Yaskawa INFORM job: 1B.JBI

/JOB
//NAME 1B
//POS
///NPOS 156,156,156,0,0,0
///TOOL 0
///POSTYPE PULSE
///PULSE
C00000=-283,-101162,-84213,3710,-80188,-1936
C00001=-283,-101162,-84213,3710,-80188,-1936
C00002=122740,19157,4035,6182,-38864,-3236
C00003=113896,2387,-35230,-12259,-73873,84724
C00004=118077,18356,-38305,-5593,-67110,82106
C00005=118077,18356,-38305,-5593,-67110,82106
C00006=124954,18047,-39669,933,-60764,50503
C00007=142043,41533,-31174,35083,-70402,26464
C00008=142043,41533,-31174,35083,-70402,26464
C00009=142043,41533,-31174,35083,-70402,26464
C00010=138380,29006,-36364,33085,-57919,16054
C00011=120169,44405,-13547,1008,-67670,-3095
C00012=105097,34464,-28801,-23051,-62948,-22596
C00013=95890,29559,-44356,-45908,-59845,-13171
C00014=95890,29559,-44356,-45908,-59845,-13171
C00015=95890,29559,-44356,-45908,-59845,-13171
C00016=100253,12469,-52865,-35215,-53568,-35172
C00017=118532,18556,-38083,-5671,-67115,-85546
C00018=114163,-2238,-37790,-11674,-74104,-76880
C00019=113860,-11716,-39905,-11456,-77647,88229
C00020=114263,6764,-46011,-12423,-64616,86905
C00021=114386,12590,-43965,-12584,-62907,81236
C00022=114386,12590,-43965,-12584,-62907,81236
C00023=125315,10262,-47133,583,-53482,49755
C00024=142444,42695,-30785,35929,-71152,26137
C00025=142444,42695,-30785,35929,-71152,26137
C00026=142444,42695,-30785,35929,-71152,26137
C00027=138388,28635,-37117,33161,-57685,15974
C00028=120215,45689,-12379,963,-68675,-3097
C00029=105043,34518,-28884,-23053,-62885,-22568
C00030=94945,31173,-44363,-48216,-61083,-12269
C00031=94945,31173,-44363,-48216,-61083,-12269
C00032=94945,31173,-44363,-48216,-61083,-12269
C00033=98921,36729,-33454,-32527,-73118,-41437
C00034=120115,8294,-47151,319,-58957,-81109
C00035=119961,110,-38118,303,-68719,-81033
C00036=104792,-5235,-37815,369,-70637,85818
C00037=99841,18984,-38422,-10534,-64752,85632
C00038=99841,18984,-38422,-10534,-64752,85632
C00039=110734,19124,-38985,1399,-60132,54528
C00040=127416,33233,-38145,36996,-63500,30231
C00041=127416,33233,-38145,36996,-63500,30231
C00042=127416,33233,-38145,36996,-63500,30231
C00043=126162,26293,-41382,40319,-54438,17642
C00044=107886,49067,-9026,3061,-69375,677
C00045=91029,44485,-19616,-23539,-67574,-17998
C00046=82208,44050,-30668,-42784,-67523,-10684
C00047=82208,44050,-30668,-42784,-67523,-10684
C00048=82208,44050,-30668,-42784,-67523,-10684
C00049=88204,44298,-22751,-24318,-76087,-40409
C00050=105281,13223,-42842,1516,-60071,-76352
C00051=104961,3103,-39460,1199,-66233,-76116
C00052=90519,4586,-31004,1943,-70415,93592
C00053=87008,29840,-27854,-8420,-66920,89435
C00054=87008,29840,-27854,-8420,-66920,89435
C00055=96155,17373,-41033,622,-52038,59586
C00056=114446,35108,-37845,43334,-60072,32327
C00057=114446,35108,-37845,43334,-60072,32327
C00058=114446,35108,-37845,43334,-60072,32327
C00059=111046,16495,-51915,50799,-38695,15495
C00060=95978,54826,-2061,4508,-68453,4441
C00061=81253,56842,-4633,-17856,-71036,-16432
C00062=73264,53266,-16777,-35142,-68308,-9926
C00063=73264,53266,-16777,-35142,-68308,-9926
C00064=73264,53266,-16777,-35142,-68308,-9926
C00065=78807,53361,-10059,-17270,-76752,-38877
C00066=91554,22306,-34303,2536,-60367,-71927
C00067=90934,11065,-29392,2410,-69140,-71537
C00068=78862,25778,-15645,3179,-69652,94598
C00069=75647,45753,-11273,-6403,-69817,92764
C00070=75647,45753,-11273,-6403,-69817,92764
C00071=83295,29982,-28891,174,-52976,64063
C00072=102305,40971,-34066,51518,-56044,33409
C00073=102305,40971,-34066,51518,-56044,33409
C00074=102305,40971,-34066,51518,-56044,33409
C00075=96997,25702,-42652,48066,-35791,21316
C00076=85385,68320,13287,6085,-70851,7845
C00077=71528,75162,16952,-15379,-76457,-14135
C00078=63937,73255,6869,-31667,-74875,-8803
C00079=63937,73255,6869,-31667,-74875,-8803
C00080=63937,73255,6869,-31667,-74875,-8803
C00081=69266,72240,11828,-14149,-81945,-36681
C00082=79459,36725,-20061,3348,-61344,-67983
C00083=78299,23264,-13932,3170,-71976,-67306
C00084=104320,15027,17892,1407,-96491,-75611
C00085=104319,15028,17890,1427,-96491,-75611
C00086=134058,-39676,-24151,-664,-98871,-85801
C00087=143372,-74915,-102054,58421,-15626,54410
C00088=139434,-25122,-70326,61306,-13879,51152
C00089=139434,-25122,-70326,61306,-13879,51152
C00090=142143,-16320,-56980,37461,-28055,41665
C00091=138227,-4635,-40701,12389,-40519,36029
C00092=135351,-979,-36711,3415,-41818,19596
C00093=134917,-12474,-49764,8729,-27792,-5734
C00094=135766,-12758,-49874,16481,-30051,-32000
C00095=132369,-15745,-53701,2097,-26646,-45047
C00096=127287,-17517,-57023,-24654,-26783,-54910
C00097=133481,-25055,-66734,-746,-13357,-86560
C00098=135802,-38388,-75052,9856,-16429,-91493
C00099=135802,-45434,-54771,5192,-32412,74887
C00100=115180,-47911,-56247,-15119,-34068,87222
C00101=119306,-82551,-105444,-10416,-9643,88947
C00102=120627,-29292,-71555,6418,-9966,79153
C00103=120627,-29292,-71555,6418,-9966,79153
C00104=125124,-22316,-61151,21013,-22926,48860
C00105=117006,-5745,-40108,-12479,-44209,48686
C00106=120091,-7318,-42638,-4085,-38918,26800
C00107=118449,-15533,-52088,-7348,-27804,5006
C00108=119516,-15941,-52128,2053,-28573,-21990
C00109=111496,-16135,-55494,-30895,-29975,-28177
C00110=111421,-17373,-56532,-32612,-31456,-48616
C00111=115167,-27509,-69100,-38565,-16380,-65993
C00112=114681,-41026,-76690,-27455,-19026,-70736
C00113=111312,-47187,-55819,-18601,-34754,89399
C00114=119856,-60423,-91419,-3428,-9742,84872
C00115=120626,-29213,-71498,6401,-9958,79150
C00116=120626,-29213,-71498,6401,-9958,79150
C00117=125772,-22206,-61200,23547,-23280,47958
C00118=126826,7414,-28064,13391,-56287,42944
C00119=120093,-7080,-42357,-4080,-38968,26798
C00120=118451,-15579,-52125,-7348,-27808,5010
C00121=119187,-16031,-52593,913,-28612,-22709
C00122=116262,-17390,-54225,-10569,-28923,-37666
C00123=104835,-15133,-61359,-62835,-35516,-38126
C00124=115015,-28488,-71572,-48615,-13974,-61504
C00125=114681,-41026,-76690,-27455,-19026,-70736
C00126=111312,-47187,-55819,-18601,-34754,89399
C00127=133743,-58056,-90173,39665,-12304,63283
C00128=131576,-28606,-72173,39560,-10330,63710
C00129=131576,-28606,-72173,39560,-10330,63710
C00130=136246,-22217,-63674,41383,-23221,46579
C00131=133839,-6410,-42313,13652,-39822,31233
C00132=135332,-14218,-52802,30045,-28779,-113
C00133=132790,-1707,-37736,16615,-42199,-13416
C00134=131751,-5560,-41359,16161,-41885,-37181
C00135=123315,-8104,-44128,-11506,-40403,-46037
C00136=118838,-21608,-64641,-49948,-24503,-46034
C00137=126445,-29920,-75490,-51443,-4984,-61687
C00138=127614,-59826,-94733,-34144,-5574,-69568
C00139=123845,-63506,-79360,-19158,-16973,85595
C00140=141900,-45604,-82921,49907,-16457,57218
C00141=140434,-25803,-72551,75363,-13806,46820
C00142=140434,-25803,-72551,75363,-13806,46820
C00143=140328,-21695,-63054,34227,-19413,40116
C00144=143522,-6973,-46080,29813,-37209,26133
C00145=141850,-4533,-42767,26469,-37315,2127
C00146=140338,-5397,-42957,25542,-37176,-18058
C00147=135954,4325,-31004,9969,-49269,-36327
C00148=127181,-6197,-43973,-18520,-39585,-44451
C00149=130222,-22519,-64075,-20467,-16747,-55259
C00150=135051,-27445,-72639,21930,-5491,-95499
C00151=139096,-69060,-94366,13448,-17195,-92631
C00152=139096,-69060,-77775,13448,-17195,71103
C00153=139096,-69060,-77775,13448,-17195,71103
C00154=-283,-101162,-84213,3710,-80188,-1936
C00155=-283,-101162,-84213,3710,-80188,-1936
BC00000=570125
BC00001=910334
BC00002=878037
BC00003=878037
BC00004=878038
BC00005=878038
BC00006=875061
BC00007=876407
BC00008=876407
BC00009=876407
BC00010=876543
BC00011=876735
BC00012=877417
BC00013=876531
BC00014=876531
BC00015=876531
BC00016=876531
BC00017=878038
BC00018=878037
BC00019=914864
BC00020=914864
BC00021=914863
BC00022=914863
BC00023=914864
BC00024=914864
BC00025=914864
BC00026=914864
BC00027=914864
BC00028=914863
BC00029=914863
BC00030=914864
BC00031=914864
BC00032=914864
BC00033=914864
BC00034=914864
BC00035=914864
BC00036=914864
BC00037=914864
BC00038=914864
BC00039=914864
BC00040=914864
BC00041=914864
BC00042=914864
BC00043=914864
BC00044=914863
BC00045=914863
BC00046=914864
BC00047=914864
BC00048=914864
BC00049=914864
BC00050=914864
BC00051=914864
BC00052=914864
BC00053=914863
BC00054=914863
BC00055=914864
BC00056=914863
BC00057=914863
BC00058=914863
BC00059=914863
BC00060=914863
BC00061=914864
BC00062=914864
BC00063=914864
BC00064=914864
BC00065=914864
BC00066=914864
BC00067=914864
BC00068=914864
BC00069=914864
BC00070=914864
BC00071=914864
BC00072=914863
BC00073=914863
BC00074=914863
BC00075=914863
BC00076=914863
BC00077=914864
BC00078=914864
BC00079=914864
BC00080=914864
BC00081=914864
BC00082=914864
BC00083=914864
BC00084=914864
BC00085=914864
BC00086=914864
BC00087=914864
BC00088=914864
BC00089=914864
BC00090=914864
BC00091=914864
BC00092=914864
BC00093=914864
BC00094=914864
BC00095=914864
BC00096=914864
BC00097=914864
BC00098=914864
BC00099=914864
BC00100=914864
BC00101=914864
BC00102=914864
BC00103=914864
BC00104=914864
BC00105=914864
BC00106=914864
BC00107=914864
BC00108=914864
BC00109=914864
BC00110=914864
BC00111=914864
BC00112=914864
BC00113=914864
BC00114=956151
BC00115=953264
BC00116=953264
BC00117=953608
BC00118=953377
BC00119=953609
BC00120=953577
BC00121=953781
BC00122=953525
BC00123=953120
BC00124=953625
BC00125=952229
BC00126=945034
BC00127=1015089
BC00128=1015089
BC00129=1015089
BC00130=1015089
BC00131=1015089
BC00132=1015089
BC00133=1015089
BC00134=1015089
BC00135=1015089
BC00136=1015089
BC00137=1015089
BC00138=1015089
BC00139=1015089
BC00140=1070064
BC00141=1070065
BC00142=1070065
BC00143=1070065
BC00144=1070065
BC00145=1070065
BC00146=1070065
BC00147=1070065
BC00148=1070065
BC00149=1070065
BC00150=1070065
BC00151=1070065
BC00152=1070065
BC00153=1070065
BC00154=1034676
BC00155=570125
EC00000=1166,0
EC00001=1166,0
EC00002=-1743,0
EC00003=-1741,0
EC00004=-1741,0
EC00005=-1741,0
EC00006=-1741,0
EC00007=-1741,0
EC00008=-1741,0
EC00009=-1741,0
EC00010=-1740,0
EC00011=-1740,0
EC00012=-1740,0
EC00013=-1740,0
EC00014=-1740,0
EC00015=-1740,0
EC00016=-1740,0
EC00017=-1741,0
EC00018=-1741,0
EC00019=-1741,0
EC00020=-1741,0
EC00021=-1741,0
EC00022=-1741,0
EC00023=-1741,0
EC00024=-1741,0
EC00025=-1741,0
EC00026=-1741,0
EC00027=-1740,0
EC00028=-1739,0
EC00029=-1740,0
EC00030=-1741,0
EC00031=-1741,0
EC00032=-1741,0
EC00033=-1740,0
EC00034=-1740,0
EC00035=-1740,0
EC00036=-1740,0
EC00037=-1740,0
EC00038=-1740,0
EC00039=-1741,0
EC00040=-1741,0
EC00041=-1741,0
EC00042=-1741,0
EC00043=-1740,0
EC00044=-1740,0
EC00045=-1740,0
EC00046=-1740,0
EC00047=-1740,0
EC00048=-1740,0
EC00049=-1740,0
EC00050=-1740,0
EC00051=-1740,0
EC00052=-1740,0
EC00053=-1741,0
EC00054=-1741,0
EC00055=-1741,0
EC00056=-1741,0
EC00057=-1741,0
EC00058=-1741,0
EC00059=-1739,0
EC00060=-1740,0
EC00061=-1740,0
EC00062=-1740,0
EC00063=-1740,0
EC00064=-1740,0
EC00065=-1740,0
EC00066=-1740,0
EC00067=-1740,0
EC00068=-1740,0
EC00069=-1741,0
EC00070=-1741,0
EC00071=-1741,0
EC00072=-1741,0
EC00073=-1741,0
EC00074=-1741,0
EC00075=-1739,0
EC00076=-1740,0
EC00077=-1740,0
EC00078=-1740,0
EC00079=-1740,0
EC00080=-1740,0
EC00081=-1740,0
EC00082=-1740,0
EC00083=-1740,0
EC00084=-1740,0
EC00085=-85617,0
EC00086=-85617,0
EC00087=-85617,0
EC00088=-85617,0
EC00089=-85617,0
EC00090=-85617,0
EC00091=-85617,0
EC00092=-85617,0
EC00093=-85617,0
EC00094=-85617,0
EC00095=-85617,0
EC00096=-85617,0
EC00097=-85617,0
EC00098=-85617,0
EC00099=-85617,0
EC00100=-85617,0
EC00101=-85617,0
EC00102=-85617,0
EC00103=-85617,0
EC00104=-85617,0
EC00105=-85617,0
EC00106=-85617,0
EC00107=-85617,0
EC00108=-85617,0
EC00109=-85617,0
EC00110=-85617,0
EC00111=-85617,0
EC00112=-85617,0
EC00113=-85617,0
EC00114=-85617,0
EC00115=-85617,0
EC00116=-85617,0
EC00117=-85617,0
EC00118=-85617,0
EC00119=-85617,0
EC00120=-85617,0
EC00121=-85617,0
EC00122=-85617,0
EC00123=-85617,0
EC00124=-85617,0
EC00125=-85617,0
EC00126=-85617,0
EC00127=-85617,0
EC00128=-85616,0
EC00129=-85616,0
EC00130=-85617,0
EC00131=-85617,0
EC00132=-85617,0
EC00133=-85617,0
EC00134=-85617,0
EC00135=-85617,0
EC00136=-85617,0
EC00137=-85617,0
EC00138=-85617,0
EC00139=-85617,0
EC00140=-85617,0
EC00141=-85617,0
EC00142=-85617,0
EC00143=-85617,0
EC00144=-85617,0
EC00145=-85617,0
EC00146=-85617,0
EC00147=-85618,0
EC00148=-85618,0
EC00149=-85618,0
EC00150=-85618,0
EC00151=-85618,0
EC00152=-85618,0
EC00153=-3792,0
EC00154=1166,0
EC00155=1166,0
//INST
///DATE 2024/12/18 10:00
///COMM OZZ
///ATTR SC,RW
///GROUP1 RB1,BS1
///GROUP2 ST1
NOP
MOVJ C00000 BC00000 VJ=70.00 DEC=20  +MOVJ EC00000 VJ=70.00
MOVJ C00001 BC00001 VJ=40.00 DEC=20  +MOVJ EC00001 VJ=0.78
MOVJ C00002 BC00002 VJ=70.00 DEC=20  +MOVJ EC00002 VJ=70.00
MOVJ C00003 BC00003 VJ=40.00 DEC=20  +MOVJ EC00003 VJ=70.00
MOVJ C00004 BC00004 VJ=40.00 DEC=20  +MOVJ EC00004 VJ=70.00
MACRO1 MJ#(0) ARGF6
ARCON
MOVC C00005 BC00005 V=5.0 DEC=20  +MOVJ EC00005 VJ=40.00
MOVC C00006 BC00006 V=5.0 DEC=20  +MOVJ EC00006 VJ=40.00
MOVC C00007 BC00007 V=5.0 DEC=20  +MOVJ EC00007 VJ=40.00
MOVJ C00008 BC00008 VJ=70.00 DEC=20  +MOVJ EC00008 VJ=40.00
MOVC C00009 BC00009 V=5.0 DEC=20  +MOVJ EC00009 VJ=40.00
MOVC C00010 BC00010 V=5.0 DEC=20  +MOVJ EC00010 VJ=40.00
MOVC C00011 BC00011 V=5.0 DEC=20  +MOVJ EC00011 VJ=40.00
MOVC C00012 BC00012 V=5.0 DEC=20  +MOVJ EC00012 VJ=40.00
MOVC C00013 BC00013 V=5.0 DEC=20  +MOVJ EC00013 VJ=40.00
MOVJ C00014 BC00014 VJ=70.00 DEC=20  +MOVJ EC00014 VJ=0.78
MOVC C00015 BC00015 V=5.0 DEC=20  +MOVJ EC00015 VJ=40.00
MOVC C00016 BC00016 V=5.0 DEC=20  +MOVJ EC00016 VJ=40.00
MOVC C00017 BC00017 V=5.0 DEC=20  +MOVJ EC00017 VJ=40.00
ARCOF
MOVJ C00018 BC00018 VJ=40.00 DEC=20  +MOVJ EC00018 VJ=40.00
MOVJ C00019 BC00019 VJ=70.00 DEC=20  +MOVJ EC00019 VJ=0.78
MOVJ C00020 BC00020 VJ=40.00 DEC=20  +MOVJ EC00020 VJ=0.78
MOVJ C00021 BC00021 VJ=40.00 DEC=20  +MOVJ EC00021 VJ=40.00
MACRO1 MJ#(0) ARGF6
ARCON
MOVC C00022 BC00022 V=5.0 DEC=20  +MOVJ EC00022 VJ=40.00
MOVC C00023 BC00023 V=5.0 DEC=20  +MOVJ EC00023 VJ=40.00
MOVC C00024 BC00024 V=5.0 DEC=20  +MOVJ EC00024 VJ=40.00
MOVJ C00025 BC00025 VJ=40.00 DEC=20  +MOVJ EC00025 VJ=40.00
MOVC C00026 BC00026 V=600.0 DEC=20  +MOVJ EC00026 VJ=40.00
MOVC C00027 BC00027 V=5.0 DEC=20  +MOVJ EC00027 VJ=40.00
MOVC C00028 BC00028 V=5.0 DEC=20  +MOVJ EC00028 VJ=40.00
MOVC C00029 BC00029 V=5.0 DEC=20  +MOVJ EC00029 VJ=40.00
MOVC C00030 BC00030 V=5.0 DEC=20  +MOVJ EC00030 VJ=40.00
MOVJ C00031 BC00031 VJ=40.00 DEC=20  +MOVJ EC00031 VJ=40.00
MOVC C00032 BC00032 V=5.0 DEC=20  +MOVJ EC00032 VJ=40.00
MOVC C00033 BC00033 V=5.0 DEC=20  +MOVJ EC00033 VJ=40.00
MOVC C00034 BC00034 V=5.0 DEC=20  +MOVJ EC00034 VJ=40.00
ARCOF
MOVJ C00035 BC00035 VJ=40.00 DEC=20  +MOVJ EC00035 VJ=40.00
MOVJ C00036 BC00036 VJ=40.00 DEC=20  +MOVJ EC00036 VJ=40.00
MOVJ C00037 BC00037 VJ=40.00 DEC=20  +MOVJ EC00037 VJ=40.00
MACRO1 MJ#(0) ARGF6
ARCON
MOVC C00038 BC00038 V=5.0 DEC=20  +MOVJ EC00038 VJ=0.78
MOVC C00039 BC00039 V=5.0 DEC=20  +MOVJ EC00039 VJ=0.78
MOVC C00040 BC00040 V=5.0 DEC=20  +MOVJ EC00040 VJ=0.78
MOVJ C00041 BC00041 VJ=40.00 DEC=20  +MOVJ EC00041 VJ=0.78
MOVC C00042 BC00042 V=600.0 DEC=20  +MOVJ EC00042 VJ=40.00
MOVC C00043 BC00043 V=5.0 DEC=20  +MOVJ EC00043 VJ=40.00
MOVC C00044 BC00044 V=5.0 DEC=20  +MOVJ EC00044 VJ=40.00
MOVC C00045 BC00045 V=5.0 DEC=20  +MOVJ EC00045 VJ=40.00
MOVC C00046 BC00046 V=5.0 DEC=20  +MOVJ EC00046 VJ=40.00
MOVJ C00047 BC00047 VJ=40.00 DEC=20  +MOVJ EC00047 VJ=40.00
MOVC C00048 BC00048 V=5.0 DEC=20  +MOVJ EC00048 VJ=40.00
MOVC C00049 BC00049 V=5.0 DEC=20  +MOVJ EC00049 VJ=40.00
MOVC C00050 BC00050 V=5.0 DEC=20  +MOVJ EC00050 VJ=40.00
ARCOF
MOVJ C00051 BC00051 VJ=40.00 DEC=20  +MOVJ EC00051 VJ=40.00
MOVJ C00052 BC00052 VJ=40.00 DEC=20  +MOVJ EC00052 VJ=40.00
MOVJ C00053 BC00053 VJ=40.00 DEC=20  +MOVJ EC00053 VJ=40.00
MACRO1 MJ#(0) ARGF6
ARCON
MOVC C00054 BC00054 V=5.0 DEC=20  +MOVJ EC00054 VJ=40.00
MOVC C00055 BC00055 V=5.0 DEC=20  +MOVJ EC00055 VJ=40.00
MOVC C00056 BC00056 V=5.0 DEC=20  +MOVJ EC00056 VJ=40.00
MOVJ C00057 BC00057 VJ=40.00 DEC=20  +MOVJ EC00057 VJ=40.00
MOVC C00058 BC00058 V=5.0 DEC=20  +MOVJ EC00058 VJ=40.00
MOVC C00059 BC00059 V=5.0 DEC=20  +MOVJ EC00059 VJ=40.00
MOVC C00060 BC00060 V=5.0 DEC=20  +MOVJ EC00060 VJ=40.00
MOVC C00061 BC00061 V=5.0 DEC=20  +MOVJ EC00061 VJ=40.00
MOVC C00062 BC00062 V=5.0 DEC=20  +MOVJ EC00062 VJ=40.00
MOVJ C00063 BC00063 VJ=40.00 DEC=20  +MOVJ EC00063 VJ=40.00
MOVC C00064 BC00064 V=5.0 DEC=20  +MOVJ EC00064 VJ=40.00
MOVC C00065 BC00065 V=5.0 DEC=20  +MOVJ EC00065 VJ=40.00
MOVC C00066 BC00066 V=5.0 DEC=20  +MOVJ EC00066 VJ=40.00
ARCOF
MOVJ C00067 BC00067 VJ=40.00 DEC=20  +MOVJ EC00067 VJ=40.00
MOVJ C00068 BC00068 VJ=40.00 DEC=20  +MOVJ EC00068 VJ=40.00
MOVJ C00069 BC00069 VJ=40.00 DEC=20  +MOVJ EC00069 VJ=40.00
MACRO1 MJ#(0) ARGF6
ARCON
MOVC C00070 BC00070 V=5.0 DEC=20  +MOVJ EC00070 VJ=40.00
MOVC C00071 BC00071 V=5.0 DEC=20  +MOVJ EC00071 VJ=40.00
MOVC C00072 BC00072 V=5.0 DEC=20  +MOVJ EC00072 VJ=40.00
MOVJ C00073 BC00073 VJ=40.00 DEC=20  +MOVJ EC00073 VJ=40.00
MOVC C00074 BC00074 V=5.0 DEC=20  +MOVJ EC00074 VJ=40.00
MOVC C00075 BC00075 V=5.0 DEC=20  +MOVJ EC00075 VJ=40.00
MOVC C00076 BC00076 V=5.0 DEC=20  +MOVJ EC00076 VJ=40.00
MOVC C00077 BC00077 V=5.0 DEC=20  +MOVJ EC00077 VJ=40.00
MOVC C00078 BC00078 V=5.0 DEC=20  +MOVJ EC00078 VJ=40.00
MOVJ C00079 BC00079 VJ=40.00 DEC=20  +MOVJ EC00079 VJ=40.00
MOVC C00080 BC00080 V=5.0 DEC=20  +MOVJ EC00080 VJ=40.00
MOVC C00081 BC00081 V=5.0 DEC=20  +MOVJ EC00081 VJ=40.00
MOVC C00082 BC00082 V=5.0 DEC=20  +MOVJ EC00082 VJ=40.00
ARCOF
MOVJ C00083 BC00083 VJ=40.00 DEC=20  +MOVJ EC00083 VJ=40.00
MOVJ C00084 BC00084 VJ=40.00 DEC=20  +MOVJ EC00084 VJ=40.00
MOVJ C00085 BC00085 VJ=40.00 DEC=20  +MOVJ EC00085 VJ=40.00
MOVJ C00086 BC00086 VJ=30.00 DEC=20  +MOVJ EC00086 VJ=30.00
MOVJ C00087 BC00087 VJ=30.00 DEC=20  +MOVJ EC00087 VJ=40.00
MOVC C00088 BC00088 V=450.0 DEC=20  +MOVJ EC00088 VJ=30.00
MACRO1 MJ#(0) ARGF6
ARCON
MOVC C00089 BC00089 V=4.7 DEC=20  +MOVJ EC00089 VJ=40.00
MOVC C00090 BC00090 V=4.7 DEC=20  +MOVJ EC00090 VJ=40.00
MOVC C00091 BC00091 V=4.7 DEC=20  +MOVJ EC00091 VJ=40.00
MOVC C00092 BC00092 V=4.7 DEC=20  +MOVJ EC00092 VJ=30.00
MOVC C00093 BC00093 V=4.2 DEC=20  +MOVJ EC00093 VJ=40.00
MOVC C00094 BC00094 V=4.2 DEC=20  +MOVJ EC00094 VJ=30.00
MOVC C00095 BC00095 V=4.2 DEC=20  +MOVJ EC00095 VJ=40.00
MOVC C00096 BC00096 V=4.2 DEC=20  +MOVJ EC00096 VJ=30.00
MOVC C00097 BC00097 V=4.2 DEC=20  +MOVJ EC00097 VJ=40.00
ARCOF
MOVJ C00098 BC00098 VJ=40.00 DEC=20  +MOVJ EC00098 VJ=40.00
MOVJ C00099 BC00099 VJ=40.00 DEC=20  +MOVJ EC00099 VJ=40.00
MOVJ C00100 BC00100 VJ=30.00 DEC=20  +MOVJ EC00100 VJ=30.00
MOVJ C00101 BC00101 VJ=30.00 DEC=20  +MOVJ EC00101 VJ=30.00
MOVC C00102 BC00102 V=450.0 DEC=20  +MOVJ EC00102 VJ=30.00
MACRO1 MJ#(0) ARGF6
ARCON
MOVC C00103 BC00103 V=5.0 DEC=20  +MOVJ EC00103 VJ=30.00
MOVC C00104 BC00104 V=5.0 DEC=20  +MOVJ EC00104 VJ=30.00
MOVC C00105 BC00105 V=5.0 DEC=20  +MOVJ EC00105 VJ=30.00
MOVC C00106 BC00106 V=5.0 DEC=20  +MOVJ EC00106 VJ=30.00
MOVC C00107 BC00107 V=5.0 DEC=20  +MOVJ EC00107 VJ=30.00
MOVC C00108 BC00108 V=5.0 DEC=20  +MOVJ EC00108 VJ=30.00
MOVC C00109 BC00109 V=5.0 DEC=20  +MOVJ EC00109 VJ=30.00
MOVC C00110 BC00110 V=5.0 DEC=20  +MOVJ EC00110 VJ=30.00
MOVC C00111 BC00111 V=5.0 DEC=20  +MOVJ EC00111 VJ=30.00
ARCOF
MOVJ C00112 BC00112 VJ=30.00 DEC=20  +MOVJ EC00112 VJ=30.00
MOVJ C00113 BC00113 VJ=30.00 DEC=20  +MOVJ EC00113 VJ=30.00
MOVJ C00114 BC00114 VJ=30.00 DEC=20  +MOVJ EC00114 VJ=0.78
MOVC C00115 BC00115 V=450.0 DEC=20  +MOVJ EC00115 VJ=30.00
ARCON
MOVC C00116 BC00116 V=5.0 DEC=20  +MOVJ EC00116 VJ=30.00
MOVC C00117 BC00117 V=5.0 DEC=20  +MOVJ EC00117 VJ=30.00
MOVC C00118 BC00118 V=5.0 DEC=20  +MOVJ EC00118 VJ=30.00
MOVC C00119 BC00119 V=5.0 DEC=20  +MOVJ EC00119 VJ=30.00
MOVC C00120 BC00120 V=5.0 DEC=20  +MOVJ EC00120 VJ=30.00
MOVC C00121 BC00121 V=5.0 DEC=20  +MOVJ EC00121 VJ=30.00
MOVC C00122 BC00122 V=5.0 DEC=20  +MOVJ EC00122 VJ=30.00
MOVC C00123 BC00123 V=5.0 DEC=20  +MOVJ EC00123 VJ=30.00
MOVC C00124 BC00124 V=5.0 DEC=20  +MOVJ EC00124 VJ=30.00
ARCOF
MOVJ C00125 BC00125 VJ=30.00 DEC=20  +MOVJ EC00125 VJ=30.00
MOVJ C00126 BC00126 VJ=30.00 DEC=20  +MOVJ EC00126 VJ=30.00
MOVJ C00127 BC00127 VJ=30.00 DEC=20  +MOVJ EC00127 VJ=30.00
MOVJ C00128 BC00128 VJ=30.00 DEC=20  +MOVJ EC00128 VJ=30.00
MACRO1 MJ#(0) ARGF6
ARCON
MOVC C00129 BC00129 V=5.0 DEC=20  +MOVJ EC00129 VJ=30.00
MOVC C00130 BC00130 V=5.0 DEC=20  +MOVJ EC00130 VJ=30.00
MOVC C00131 BC00131 V=5.0 DEC=20  +MOVJ EC00131 VJ=30.00
MOVC C00132 BC00132 V=5.0 DEC=20  +MOVJ EC00132 VJ=30.00
MOVC C00133 BC00133 V=5.0 DEC=20  +MOVJ EC00133 VJ=30.00
MOVC C00134 BC00134 V=5.0 DEC=20  +MOVJ EC00134 VJ=30.00
MOVC C00135 BC00135 V=5.0 DEC=20  +MOVJ EC00135 VJ=30.00
MOVC C00136 BC00136 V=5.0 DEC=20  +MOVJ EC00136 VJ=30.00
MOVC C00137 BC00137 V=5.0 DEC=20  +MOVJ EC00137 VJ=30.00
ARCOF
MOVJ C00138 BC00138 VJ=30.00 DEC=20  +MOVJ EC00138 VJ=30.00
MOVJ C00139 BC00139 VJ=30.00 DEC=20  +MOVJ EC00139 VJ=30.00
MOVJ C00140 BC00140 VJ=30.00 DEC=20  +MOVJ EC00140 VJ=30.00
MOVJ C00141 BC00141 VJ=30.00 DEC=20  +MOVJ EC00141 VJ=30.00
MACRO1 MJ#(0) ARGF6
ARCON
MOVC C00142 BC00142 V=5.0 DEC=20  +MOVJ EC00142 VJ=30.00
MOVC C00143 BC00143 V=5.0 DEC=20  +MOVJ EC00143 VJ=30.00
MOVC C00144 BC00144 V=5.0 DEC=20  +MOVJ EC00144 VJ=30.00
MOVC C00145 BC00145 V=5.0 DEC=20  +MOVJ EC00145 VJ=30.00
MOVC C00146 BC00146 V=5.0 DEC=20  +MOVJ EC00146 VJ=30.00
MOVC C00147 BC00147 V=5.0 DEC=20  +MOVJ EC00147 VJ=30.00
MOVC C00148 BC00148 V=5.0 DEC=20  +MOVJ EC00148 VJ=30.00
MOVC C00149 BC00149 V=5.0 DEC=20  +MOVJ EC00149 VJ=30.00
MOVC C00150 BC00150 V=5.0 DEC=20  +MOVJ EC00150 VJ=30.00
ARCOF
MOVJ C00151 BC00151 VJ=30.00 DEC=20  +MOVJ EC00151 VJ=30.00
MOVJ C00152 BC00152 VJ=30.00 DEC=20  +MOVJ EC00152 VJ=30.00
MOVJ C00153 BC00153 VJ=30.00 DEC=20  +MOVJ EC00153 VJ=30.00
MOVJ C00154 BC00154 VJ=40.00 DEC=20  +MOVJ EC00154 VJ=40.00
MOVJ C00155 BC00155 VJ=40.00 DEC=20  +MOVJ EC00155 VJ=40.00
END
